(* IEC 61131-3 sources: rusty/tests/lit/multi/library_string_overflow, 1 file *)

(* ---- library_string_overflow_prog.st ---- *)
FUNCTION main
VAR
    MyString : STRING;
    MyInt : INT := 1234;
    MyGuard : DINT := 24681357;
    retValue : ErrorCode;
END_VAR

retValue := Config_GetString('/service/config/logLevel', MyString);
printf('ret=%d my_int=%d my_guard=%d value_prefix=%.8s', retValue, MyInt, MyGuard, MyString);
// CHECK: ret=0 my_int=1234 my_guard=24681357 value_prefix=AAAAAAAA
END_FUNCTION
